FUNCTION_BLOCK FB_ReactorValves_Test EXTENDS TcUnit.FB_TestSuite
VAR_INPUT
END_VAR
VAR_OUTPUT
END_VAR
VAR
END_VAR


// Valve should open if upper interval reached
valveShouldOpenIfUpperIntervalReached();

METHOD valveShouldCloseIfForcedTo
VAR
	valves : FB_ReactorValves;
END_VAR

TEST('valve Should close if forced to');
			
	valves.pressureIntervalControl(
		interval_1_condition:= TRUE, 
		pressureUpperInterval_1:= 20, 
		pressureLowerInterval_1:= 0, 
		interval_2_condition:= FALSE, 
		pressureUpperInterval_2:= 999, 
		pressureLowerInterval_2:= 999, 
		interval_3_condition:= FALSE, 
		pressureUpperInterval_3:= 999, 
		pressureLowerInterval_3:= 999, 
		pressureValue:= 220, 
		pressureReference:= 200, 
		valveOpenCondition:= FALSE, 
		forceValveClosed:= FALSE);
			
	AssertEquals_BOOL(Expected :=  FALSE, Actual := valves.pressureControlOpen, Message := 'Valve not closed when forced to');	
TEST_FINISHED();
END_METHOD

METHOD valveShouldCloseIfLowerIntervalReached
VAR
	valves : FB_ReactorValves;
END_VAR

TEST('valve Should Close If Lower Interval Reached');
			
	valves.pressureIntervalControl(
		interval_1_condition:= TRUE, 
		pressureUpperInterval_1:= 20, 
		pressureLowerInterval_1:= 0, 
		interval_2_condition:= FALSE, 
		pressureUpperInterval_2:= 999, 
		pressureLowerInterval_2:= 999, 
		interval_3_condition:= FALSE, 
		pressureUpperInterval_3:= 999, 
		pressureLowerInterval_3:= 999, 
		pressureValue:= 220, 
		pressureReference:= 200, 
		valveOpenCondition:= TRUE, 
		forceValveClosed:= FALSE);
		
	valves.pressureIntervalControl(
		interval_1_condition:= TRUE, 
		pressureUpperInterval_1:= 20, 
		pressureLowerInterval_1:= 20, 
		interval_2_condition:= FALSE, 
		pressureUpperInterval_2:= 999, 
		pressureLowerInterval_2:= 999, 
		interval_3_condition:= FALSE, 
		pressureUpperInterval_3:= 999, 
		pressureLowerInterval_3:= 999, 
		pressureValue:= 180, 
		pressureReference:= 200, 
		valveOpenCondition:= TRUE, 
		forceValveClosed:= FALSE);
			
	AssertEquals_BOOL(Expected :=  FALSE, Actual := valves.pressureControlOpen, Message := 'Valve not closed when lower interval reached');	
TEST_FINISHED();
END_METHOD

METHOD valveShouldCloseIfOpenConditionNotFulfilled
VAR
	valves : FB_ReactorValves;
END_VAR

TEST('valve Should close if open condition not fulfilled');
			
	valves.pressureIntervalControl(
		interval_1_condition:= TRUE, 
		pressureUpperInterval_1:= 20, 
		pressureLowerInterval_1:= 0, 
		interval_2_condition:= FALSE, 
		pressureUpperInterval_2:= 999, 
		pressureLowerInterval_2:= 999, 
		interval_3_condition:= FALSE, 
		pressureUpperInterval_3:= 999, 
		pressureLowerInterval_3:= 999, 
		pressureValue:= 220, 
		pressureReference:= 200, 
		valveOpenCondition:= FALSE, 
		forceValveClosed:= FALSE);
			
	AssertEquals_BOOL(Expected :=  FALSE, Actual := valves.pressureControlOpen, Message := 'Valve not closed when open condition not fulfilled');	
TEST_FINISHED();
END_METHOD

METHOD valveShouldOpenIfUpperIntervalReached
VAR
	valves : FB_ReactorValves;
END_VAR

TEST('valve Should Open If Upper Interval Reached');
			
	valves.pressureIntervalControl(
		interval_1_condition:= TRUE, 
		pressureUpperInterval_1:= 20, 
		pressureLowerInterval_1:= 0, 
		interval_2_condition:= FALSE, 
		pressureUpperInterval_2:= 999, 
		pressureLowerInterval_2:= 999, 
		interval_3_condition:= FALSE, 
		pressureUpperInterval_3:= 999, 
		pressureLowerInterval_3:= 999, 
		pressureValue:= 220, 
		pressureReference:= 200, 
		valveOpenCondition:= TRUE, 
		forceValveClosed:= FALSE);
			
	AssertEquals_BOOL(Expected :=  TRUE, Actual := valves.pressureControlOpen, Message := 'Valve not opened when upper interval reached');	
TEST_FINISHED();
END_METHOD

END_FUNCTION_BLOCK

(* stored: Version 1.1.0.1, ProductVersion 3.1.4024.9
   POU FB_ReactorValves_Test: Id {eb6e6a1a-c546-4e6a-9c45-f02a2bb7f3d2}, SpecialFunc None
   Method valveShouldCloseIfForcedTo: Id {f4be1906-027b-48de-af99-f6d33283511b}
   Method valveShouldCloseIfLowerIntervalReached: Id {8342c621-d981-480d-9d63-1f2522286490}
   Method valveShouldCloseIfOpenConditionNotFulfilled: Id {e2b33ad6-0094-45e0-949f-42107b8a50cd}
   Method valveShouldOpenIfUpperIntervalReached: Id {2e665aa1-ec34-4395-9c56-38bd77bd1367} *)
